(* IEC 61131-3 sources: rusty/tests/lit/multi/interface_consumer_separate_file, 4 files *)

(* ---- iface.st ---- *)
INTERFACE IFoo
    METHOD bar : DINT
    END_METHOD
END_INTERFACE

(* ---- main.st ---- *)
FUNCTION main
    VAR
        impl : FbImpl;
        consumer : FbConsumer;
    END_VAR

    consumer.setRef(impl);
    printf('%d$N', consumer.invoke());
END_FUNCTION

(* ---- consumer.st ---- *)
FUNCTION_BLOCK FbConsumer
    VAR
        stored : IFoo;
    END_VAR

    METHOD setRef
        VAR_INPUT
            iface : IFoo;
        END_VAR
        stored := iface;
    END_METHOD

    METHOD invoke : DINT
        invoke := stored.bar();
    END_METHOD
END_FUNCTION_BLOCK

(* ---- impl.st ---- *)
FUNCTION_BLOCK FbImpl IMPLEMENTS IFoo
    METHOD bar : DINT
        bar := 42;
    END_METHOD
END_FUNCTION_BLOCK
